(* PLC project TBEN_L5_PLC11.project, CODESYS CODESYS V3.5 SP21 Patch 1 *)
(* stored: creationDateTime 2026-11-07T15:35:08.2741952, modificationDateTime 2026-11-07T15:09:07.4034196 *)

// Đọc Float32T IO-Link (IEEE754 big-endian): chép bit pattern, không đổi số học
FUNCTION F_IolGetR32BE : REAL
VAR_INPUT
    pBuf  : POINTER TO BYTE;
    uiOff : UINT;
END_VAR
VAR
    dwTmp : DWORD;
    pR    : POINTER TO REAL;
END_VAR

            dwTmp := F_IolGetU32BE(pBuf, uiOff);
pR := ADR(dwTmp);
F_IolGetR32BE := pR^;

          
END_FUNCTION
